(* IEC 61131-3 sources: llm-plc-st-eval/data/processed_v2/claude-sonnet-4-6/B5/few_shot, 3 files *)

(* ---- ejec_1.st ---- *)
FUNCTION_BLOCK FB_Ventilador
VAR_INPUT
    quemadorOn : BOOL; (* Señal del quemador: TRUE = encendido *)
END_VAR
VAR_OUTPUT
    ventilador : BOOL; (* Salida del ventilador de enfriamiento *)
END_VAR
VAR
    tPostMarcha : TON; (* Temporizador de post-marcha *)
END_VAR

(* El temporizador arranca cuando el quemador se apaga (flanco descendente) *)
(* IN = FALSE detiene/resetea el timer; IN = TRUE lo pone en marcha         *)
tPostMarcha(IN := NOT quemadorOn, PT := T#30S);

(* El ventilador funciona mientras el quemador este encendido               *)
(* o mientras el temporizador de post-marcha no haya concluido              *)
ventilador := quemadorOn OR NOT tPostMarcha.Q;
END_FUNCTION_BLOCK

(* ---- ejec_2.st ---- *)
FUNCTION_BLOCK FB_Ventilador
VAR_INPUT
    quemadorOn : BOOL; (* Señal del quemador: TRUE = encendido *)
END_VAR
VAR_OUTPUT
    ventilador : BOOL; (* Salida del ventilador de enfriamiento *)
END_VAR
VAR
    tPostMarcha : TOF; (* Temporizador de retardo a la desconexion *)
END_VAR

(* El ventilador funciona mientras el quemador este encendido         *)
(* y continua 30 s adicionales tras apagarse el quemador (post-marcha) *)
tPostMarcha(IN := quemadorOn, PT := T#30S);
ventilador := tPostMarcha.Q;
END_FUNCTION_BLOCK

(* ---- ejec_3.st ---- *)
FUNCTION_BLOCK FB_Ventilador
VAR_INPUT
    quemadorOn : BOOL; (* Señal del quemador: TRUE = encendido *)
END_VAR
VAR_OUTPUT
    ventilador : BOOL; (* Salida del ventilador de enfriamiento *)
END_VAR
VAR
    tPostMarcha : TOF; (* Temporizador de retardo a la desconexion *)
END_VAR

(* El ventilador funciona mientras el quemador este encendido        *)
(* y continua 30 s adicionales tras apagarse el quemador (post-marcha) *)
tPostMarcha(IN := quemadorOn, PT := T#30S);
ventilador := tPostMarcha.Q;
END_FUNCTION_BLOCK
